Fanuc KAREL source: kb00116.KL

PROGRAM KB00116
%NOLOCKGROUP
VAR
P1:REAL;RESULT:REAL
BEGIN
--
P1=1.0
RESULT=LN(P1)
END KB00116
